Yaskawa INFORM job: R1-HOME.JBI

/JOB
//NAME R1-HOME
//POS
///NPOS 0,0,0,1,0,0
///TOOL 0
///POSTYPE PULSE
///PULSE
P00100=-3000,48000,-36000,0,-95000,0
//INST
///DATE 2023/11/01 07:45
///ATTR SC,RW
///GROUP1 RB1
NOP
MOVJ P100 VJ=25.00
END
